Fanuc KAREL source: ko00078.KL

-- PROVISIONAL review KL for V1013-1; original PC SHA256 73e41096ab0020cff13dfb041a265cfa9f655694dddc951df99201eddc9f56af
-- Incomplete behavior may be omitted. Consult companion uncertainty JSON. Do not deploy.
PROGRAM KO00078
%NOLOCKGROUP
BEGIN
  -- UNRESOLVED_PC offsets 5-12; opcodes 9D,23
  -- UNRESOLVED_PC offsets 17-66; opcodes 27,22,1C,27,49,7E,AD,22,31,7E,4A
  -- UNRESOLVED_PC offsets 71-75; opcodes 7F
END KO00078
